INTERFACE I_UnitLimitRule EXTENDS I_Module

METHOD M_Evaluate : ST_LimitOut	// 유닛 P·Q 한도 (사용자 한도 등). bActive = FALSE면 제한 없음. 범위를 좁히기만 함 (0은 항상 허용)
VAR_INPUT
	i_stView	: ST_UnitLimitView;
END_VAR
END_METHOD

END_INTERFACE

(* stored: Version 1.1.0.1, ProductVersion 3.1.4024.15
   Itf I_UnitLimitRule: Id {40addec0-30c6-43a7-9c84-d8d611ecf8c5}
   Method M_Evaluate: Id {4b4a50f7-ffc1-4881-ae6d-9093336fe5f8} *)
